{region 'Documentation'}
(*!
<summary>Check that IN is at most Maximum.</summary>
*)
{endregion}
FUNCTION_BLOCK AssertLessEqual_LInt EXTENDS AssertionBase
VAR_INPUT
    IN : LINT; //! Actual value checked or observed by this Assertion.
    Maximum : LINT; //! Inclusive upper bound of the comparison; for a range, must not be below Minimum.
END_VAR

SUPER^();

{region 'Documentation'}
(*!
<summary>Check that IN is at most Maximum.</summary>
*)
{endregion}
METHOD PROTECTED Assert
VAR
    Message : STRING(GVL_Constants.MessageLength);
    MaximumText : STRING(GVL_Constants.AssertionValueLength);
    ActualText : STRING(GVL_Constants.AssertionValueLength);
END_VAR
IF NOT EvaluationActive THEN
    RETURN;
END_IF;

IF Result = E_Result.Error THEN
    RETURN;
END_IF;

IF Result = E_Result.Failed THEN
    RETURN;
END_IF;

IF IN > Maximum THEN
    MaximumText := LINT_TO_STRING(Maximum);
    ActualText := LINT_TO_STRING(IN);
    Message := CONCAT('Assertion failed: value is above maximum. Maximum = ',
        MaximumText);
    Message := CONCAT(Message, ', Actual = ');
    Message := CONCAT(Message, ActualText);
    Message := CONCAT(Message, '.');
    Fail(Message := Message);
    RETURN;
END_IF;

Pass();
END_METHOD

END_FUNCTION_BLOCK

(* stored: Version 1.1.0.1
   POU AssertLessEqual_LInt: Id {de5093be-701f-4b78-9cab-669433b95029}, SpecialFunc None
   Folder Internal: Id {9f31eaae-d7d6-43a5-96f1-286902f5fd0a}
   Method Assert: Id {2485fb33-bbf1-4ca2-9ab2-38941d884f6c} *)
